Fanuc KAREL source: KT00527.KL

PROGRAM KT00527
%NOLOCKGROUP
VAR
  P1: XYZWPREXT
  P2: XYZWPREXT
  OUT: JOINTPOS
BEGIN
  P1.X = 1.0
  P2.Y = 2.0
  P1.X = 1.0
  P2.Y = 2.0
  OUT = P1 : P2
END KT00527
